FUNCTION_BLOCK FB_HeaterPI (* Migrated from IEC 61131-3 ST *)
  (* Standard: 61499-2 *)
  (* Version 1.0, 2026-11-06, st2fb *)
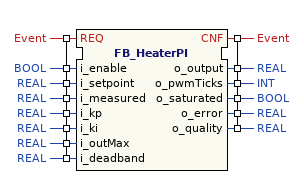
  EVENT_INPUT
    REQ WITH i_enable, i_setpoint, i_measured, i_kp, i_ki, i_outMax, i_deadband;
  END_EVENT
  EVENT_OUTPUT
    CNF WITH o_output, o_pwmTicks, o_saturated, o_error, o_quality;
  END_EVENT
  VAR_INPUT
    i_enable : BOOL;
    i_setpoint : REAL;
    i_measured : REAL;
    i_kp : REAL;
    i_ki : REAL;
    i_outMax : REAL;
    i_deadband : REAL;
  END_VAR
  VAR_OUTPUT
    o_output : REAL;
    o_pwmTicks : INT;
    o_saturated : BOOL;
    o_error : REAL;
    o_quality : REAL;
  END_VAR
  VAR
    statIntegral : REAL := 0.0;
    statFirstRun : BOOL := TRUE;
    tempUnclamped : REAL := 0.0;
    tempErrorAbs : REAL := 0.0;
  END_VAR
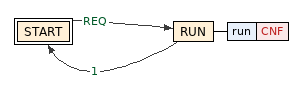
  EC_STATES
    START;
    RUN : run -> CNF;
  END_STATES
  EC_TRANSITIONS
    START TO RUN := REQ;
    RUN TO START := 1;
  END_TRANSITIONS
  ALGORITHM run IN ST:
IF NOT i_enable THEN
  o_saturated := FALSE;
  statFirstRun := TRUE;
ELSE
  IF statFirstRun THEN
    statIntegral := o_output;
    statFirstRun := FALSE;
  END_IF;
  o_error := i_setpoint - i_measured;
  tempErrorAbs := ABS(o_error);
  IF tempErrorAbs < i_deadband THEN
    o_error := 0.0;
  END_IF;
  tempUnclamped := i_kp * o_error + statIntegral + i_ki * o_error;
  o_output := LIMIT(0.0, tempUnclamped, i_outMax);
  o_saturated := o_output <> tempUnclamped;
  IF NOT o_saturated THEN
    statIntegral := statIntegral + i_ki * o_error;
  END_IF;
  o_pwmTicks := DINT_TO_INT(REAL_TO_DINT(o_output * 10.0));
  o_quality := SQRT(o_error * o_error + 1.0);
END_IF;
  END_ALGORITHM
END_FUNCTION_BLOCK
